// I_Comm stub that records the Publish* calls of a test (parameter name, kind, value), for the telemetry characterization
// (IagTelemetry_Tests). Like FB_NullComm every call reports success. Recording is off until Start(), so the suites that
// do not look at the telemetry pay only the memory.
// Kinds: 1 LREAL, 2 INT (value as LREAL), 3 BOOL (0.0/1.0), 4 STRING (value not kept), 5 Publish (not kept).
FUNCTION_BLOCK FB_RecordingComm IMPLEMENTS BROTLib.I_Comm
VAR_OUTPUT
	nCount		: INT;			// records in aNames/aKinds/aValues (1..nCount)
	bOverflow	: BOOL;			// more than 160 calls: the last slot holds the newest call
	aNames		: ARRAY[1..160] OF STRING(80);
	aKinds		: ARRAY[1..160] OF INT;
	aValues		: ARRAY[1..160] OF LREAL;
END_VAR
VAR
	bRecording	: BOOL;
	sFilter		: STRING(80);
END_VAR

METHOD Publish : BOOL
VAR_INPUT
	domain			: STRING(255) := 'environment';
	location		: STRING(255) := 'roof';
	parameter		: STRING(255);
	value			: STRING(255);
END_VAR
VAR_OUTPUT
	published	: BOOL;
END_VAR
Record(sName := parameter, nKind := 5, fValue := 0.0);
Publish := TRUE;
published := TRUE;
END_METHOD

METHOD PublishLREAL : BOOL
VAR_INPUT
	domain			: STRING(255) := 'environment';
	location		: STRING(255) := 'roof';
	parameter		: STRING(255);
	value			: LREAL;
END_VAR
VAR_OUTPUT
	published	: BOOL;
END_VAR
Record(sName := parameter, nKind := 1, fValue := value);
PublishLREAL := TRUE;
published := TRUE;
END_METHOD

METHOD PublishINT : BOOL
VAR_INPUT
	domain			: STRING(255) := 'environment';
	location		: STRING(255) := 'roof';
	parameter		: STRING(255);
	value			: LINT;
END_VAR
VAR_OUTPUT
	published	: BOOL;
END_VAR
Record(sName := parameter, nKind := 2, fValue := LINT_TO_LREAL(value));
PublishINT := TRUE;
published := TRUE;
END_METHOD

METHOD PublishBOOL : BOOL
VAR_INPUT
	domain			: STRING(255) := 'environment';
	location		: STRING(255) := 'roof';
	parameter		: STRING(255);
	value			: BOOL;
END_VAR
VAR_OUTPUT
	published	: BOOL;
END_VAR
Record(sName := parameter, nKind := 3, fValue := SEL(value, 0.0, 1.0));
PublishBOOL := TRUE;
published := TRUE;
END_METHOD

METHOD PublishString : BOOL
VAR_INPUT
	domain			: STRING(255) := 'environment';
	location		: STRING(255) := 'roof';
	parameter		: STRING(255);
	value			: STRING(255);
END_VAR
VAR_OUTPUT
	published	: BOOL;
END_VAR
Record(sName := parameter, nKind := 4, fValue := 0.0);
PublishString := TRUE;
published := TRUE;
END_METHOD

METHOD PublishLog : BOOL
VAR_INPUT
	level		: STRING(255) := 'INFO';
	message		: STRING(255);
END_VAR
VAR_OUTPUT
	published	: BOOL;
END_VAR
PublishLog := TRUE;
published := TRUE;
END_METHOD

METHOD PRIVATE Record
VAR_INPUT
	sName	: STRING(255);
	nKind	: INT;
	fValue	: LREAL;
END_VAR
VAR
	nIndex	: INT;
END_VAR
IF NOT bRecording THEN
	RETURN;
END_IF
IF sFilter <> '' AND sFilter <> sName THEN
	RETURN;
END_IF
IF nCount >= 160 THEN
	// full: the last slot keeps the latest call, so a filtered recording still ends with the newest value
	bOverflow := TRUE;
	nIndex := 160;
ELSE
	nCount := nCount + 1;
	nIndex := nCount;
END_IF
aNames[nIndex] := sName;
aKinds[nIndex] := nKind;
aValues[nIndex] := fValue;
END_METHOD

// Clears the record and starts recording; sNameFilter <> '' records only calls with that parameter name.
METHOD Start
VAR_INPUT
	sNameFilter	: STRING(80);
END_VAR
VAR
	i	: INT;
END_VAR
FOR i := 1 TO 160 DO
	aNames[i] := '';
	aKinds[i] := 0;
	aValues[i] := 0.0;
END_FOR
nCount := 0;
bOverflow := FALSE;
sFilter := sNameFilter;
bRecording := TRUE;
END_METHOD

METHOD Stop
bRecording := FALSE;
END_METHOD

// first record with this parameter name, 0 if none
METHOD FindName : INT
VAR_INPUT
	sName	: STRING(80);
END_VAR
VAR
	i	: INT;
END_VAR
FindName := 0;
FOR i := 1 TO nCount DO
	IF aNames[i] = sName THEN
		FindName := i;
		RETURN;
	END_IF
END_FOR
END_METHOD

END_FUNCTION_BLOCK

(* stored: Version 1.1.0.1, ProductVersion 3.1.4024.15
   POU FB_RecordingComm: Id {16e8d6e3-62c4-4300-b64b-3dddd69dc399}, SpecialFunc None
   Method Publish: Id {d09c4159-f8aa-400f-be89-f06f0ddd0a4a}
   Method PublishLREAL: Id {455f469c-4b43-4249-896f-d7439b51c2c5}
   Method PublishINT: Id {ec3142d8-e5ea-4779-aa0b-4ef06ffa9c51}
   Method PublishBOOL: Id {8aecab3e-bd9d-48e3-8165-b7d92bebd1d5}
   Method PublishString: Id {05a26dcd-a3b8-4a40-a81c-bc8e3af7bb52}
   Method PublishLog: Id {6ba5f234-0740-44d5-8971-260f7df4f23a}
   Method Record: Id {c242eb64-765d-4bf2-b5a7-6ed49034b742}
   Method Start: Id {5af6e0a8-b4c6-411c-a029-00684622728b}
   Method Stop: Id {e2e8b470-f139-4271-8923-62aa6ed0aac3}
   Method FindName: Id {9e9ccefe-b5e0-4803-af39-8b7116da0597} *)
